(* IEC 61131-3 sources: sis-interlock-demo/tests/GVLs/Generated, 2 files *)

(* ---- GVL_TestsGenerated.gvl.st ---- *)
// AUTO-GENERATED by cemgen 1.0.0 — не редактировать: правьте матрицу и запустите
//   python -m cemgen generate <файл матрицы .csv или .xlsx>
// Матрица: SIS-V101-CEM, объект V-101, ревизия B от 2026-10-19, SHA-256 сетки df2ed4841a9453ca
// Назначение: экземпляры сгенерированных наборов coUnit: таблицы истинности голосования и сценарии
//             по матрице. {attribute 'linkalways'} обязателен: без него CODESYS выбрасывает GVL, на
//             которую никто не ссылается, и наборы молча пропадают.
// Автор:      kr0nsch; код — генератор cemgen
// Версия:     1.0.0
// Документ:   docs/DESIGN.md, раздел «10. Генератор cemgen»; docs/cause_effect_matrix.md
// ВНИМАНИЕ:   код демонстрационный и не предназначен для систем безопасности. Реальная ПАЗ требует
//             определения SIL, сертифицированных аппаратных и программных средств и валидации по
//             ГОСТ Р МЭК 61511.
{attribute 'qualified_only'}
{attribute 'linkalways'}
VAR_GLOBAL
    fbVoteTruthTest : FB_VoteTruth_Test;   // таблицы истинности голосования (36 тестов)
    fbCemGen01Test  : FB_CemGen01_Test;    // сценарии по матрице, тесты 1–40
    fbCemGen02Test  : FB_CemGen02_Test;    // сценарии по матрице, тесты 41–80
    fbCemGen03Test  : FB_CemGen03_Test;    // сценарии по матрице, тесты 81–83
END_VAR

(* ---- GVL_VoteTruthTable.gvl.st ---- *)
// AUTO-GENERATED by cemgen 1.0.0 — не редактировать: правьте матрицу и запустите
//   python -m cemgen generate <файл матрицы .csv или .xlsx>
// Матрица: SIS-V101-CEM, объект V-101, ревизия B от 2026-10-19, SHA-256 сетки df2ed4841a9453ca
// Назначение: таблицы истинности голосования (DESIGN.md, 12.2): ожидаемые байты результата
//             F_VoteEval (уровень 1) и FB_Voting (уровень 2) для всех схем, политик и видов входа;
//             считает эталонная модель cemgen. Байт: бит 0 — xTrip, бит 1 — xDegraded, биты 2–4 —
//             eArchEff (0 None, 1 1oo1, 2 1oo2, 3 2oo2, 4 2oo3, 5 ForcedTrip), биты 5–7 — байпас
//             каналов 1–3 Active (уровень 2).
// Автор:      kr0nsch; код — генератор cemgen
// Версия:     1.0.0
// Документ:   docs/DESIGN.md, раздел «10. Генератор cemgen»; docs/cause_effect_matrix.md
// ВНИМАНИЕ:   код демонстрационный и не предназначен для систем безопасности. Реальная ПАЗ требует
//             определения SIL, сертифицированных аппаратных и программных средств и валидации по
//             ГОСТ Р МЭК 61511.
{attribute 'qualified_only'}
VAR_GLOBAL CONSTANT
    // Уровень 1 — F_VoteEval: строка r, состояние канала k — (r SHR 2(k − 1)) AND 3:
    // 0 Normal, 1 Demand, 2 Invalid, 3 Bypassed; каналы k > N — NotUsed
    TT_EVAL_1OO1_VT : ARRAY[0..3] OF BYTE := [
        16#04, 16#05, 16#17, 16#17];
    TT_EVAL_1OO1_DS : ARRAY[0..3] OF BYTE := [
        16#04, 16#05, 16#17, 16#17];
    TT_EVAL_1OO1_DA : ARRAY[0..3] OF BYTE := [
        16#04, 16#05, 16#17, 16#17];
    TT_EVAL_1OO2_VT : ARRAY[0..15] OF BYTE := [
        16#08, 16#09, 16#17, 16#06, 16#09, 16#09, 16#17, 16#07, 16#17, 16#17, 16#17, 16#17, 16#06, 16#07, 16#17, 16#17];
    TT_EVAL_1OO2_DS : ARRAY[0..15] OF BYTE := [
        16#08, 16#09, 16#06, 16#06, 16#09, 16#09, 16#07, 16#07, 16#06, 16#07, 16#17, 16#17, 16#06, 16#07, 16#17, 16#17];
    TT_EVAL_1OO2_DA : ARRAY[0..15] OF BYTE := [
        16#08, 16#09, 16#06, 16#06, 16#09, 16#09, 16#07, 16#07, 16#06, 16#07, 16#17, 16#17, 16#06, 16#07, 16#17, 16#17];
    TT_EVAL_2OO2_VT : ARRAY[0..15] OF BYTE := [
        16#0C, 16#0C, 16#06, 16#06, 16#0C, 16#0D, 16#07, 16#07, 16#06, 16#07, 16#17, 16#17, 16#06, 16#07, 16#17, 16#17];
    TT_EVAL_2OO2_DS : ARRAY[0..15] OF BYTE := [
        16#0C, 16#0C, 16#06, 16#06, 16#0C, 16#0D, 16#07, 16#07, 16#06, 16#07, 16#17, 16#17, 16#06, 16#07, 16#17, 16#17];
    TT_EVAL_2OO2_DA : ARRAY[0..15] OF BYTE := [
        16#0C, 16#0C, 16#06, 16#06, 16#0C, 16#0D, 16#07, 16#07, 16#06, 16#07, 16#17, 16#17, 16#06, 16#07, 16#17, 16#17];
    TT_EVAL_2OO3_VT : ARRAY[0..63] OF BYTE := [
        16#10, 16#10, 16#0A, 16#0A, 16#10, 16#11, 16#0B, 16#0B, 16#0A, 16#0B, 16#17, 16#17, 16#0A, 16#0B, 16#17, 16#06,
        16#10, 16#11, 16#0B, 16#0B, 16#11, 16#11, 16#0B, 16#0B, 16#0B, 16#0B, 16#17, 16#17, 16#0B, 16#0B, 16#17, 16#07,
        16#0A, 16#0B, 16#17, 16#17, 16#0B, 16#0B, 16#17, 16#17, 16#17, 16#17, 16#17, 16#17, 16#17, 16#17, 16#17, 16#17,
        16#0A, 16#0B, 16#17, 16#06, 16#0B, 16#0B, 16#17, 16#07, 16#17, 16#17, 16#17, 16#17, 16#06, 16#07, 16#17, 16#17];
    TT_EVAL_2OO3_DS : ARRAY[0..63] OF BYTE := [
        16#10, 16#10, 16#0A, 16#0A, 16#10, 16#11, 16#0B, 16#0B, 16#0A, 16#0B, 16#06, 16#06, 16#0A, 16#0B, 16#06, 16#06,
        16#10, 16#11, 16#0B, 16#0B, 16#11, 16#11, 16#0B, 16#0B, 16#0B, 16#0B, 16#07, 16#07, 16#0B, 16#0B, 16#07, 16#07,
        16#0A, 16#0B, 16#06, 16#06, 16#0B, 16#0B, 16#07, 16#07, 16#06, 16#07, 16#17, 16#17, 16#06, 16#07, 16#17, 16#17,
        16#0A, 16#0B, 16#06, 16#06, 16#0B, 16#0B, 16#07, 16#07, 16#06, 16#07, 16#17, 16#17, 16#06, 16#07, 16#17, 16#17];
    TT_EVAL_2OO3_DA : ARRAY[0..63] OF BYTE := [
        16#10, 16#10, 16#0E, 16#0E, 16#10, 16#11, 16#0E, 16#0E, 16#0E, 16#0E, 16#06, 16#06, 16#0E, 16#0E, 16#06, 16#06,
        16#10, 16#11, 16#0E, 16#0E, 16#11, 16#11, 16#0F, 16#0F, 16#0E, 16#0F, 16#07, 16#07, 16#0E, 16#0F, 16#07, 16#07,
        16#0E, 16#0E, 16#06, 16#06, 16#0E, 16#0F, 16#07, 16#07, 16#06, 16#07, 16#17, 16#17, 16#06, 16#07, 16#17, 16#17,
        16#0E, 16#0E, 16#06, 16#06, 16#0E, 16#0F, 16#07, 16#07, 16#06, 16#07, 16#17, 16#17, 16#06, 16#07, 16#17, 16#17];
    // Уровень 2 — FB_Voting: строка r, биты канала k — 3(k − 1): требование, достоверность,
    // запрос байпаса; на строку два вызова одного экземпляра (сначала без запросов байпаса)
    TT_FB_1OO1_VT_DI : ARRAY[0..7] OF BYTE := [
        16#17, 16#17, 16#04, 16#05, 16#17, 16#17, 16#04, 16#05];
    TT_FB_1OO1_VT_AI : ARRAY[0..7] OF BYTE := [
        16#17, 16#17, 16#04, 16#05, 16#17, 16#17, 16#04, 16#05];
    TT_FB_1OO1_DS_DI : ARRAY[0..7] OF BYTE := [
        16#17, 16#17, 16#04, 16#05, 16#17, 16#17, 16#04, 16#05];
    TT_FB_1OO1_DS_AI : ARRAY[0..7] OF BYTE := [
        16#17, 16#17, 16#04, 16#05, 16#17, 16#17, 16#04, 16#05];
    TT_FB_1OO1_DA_DI : ARRAY[0..7] OF BYTE := [
        16#17, 16#17, 16#04, 16#05, 16#17, 16#17, 16#04, 16#05];
    TT_FB_1OO1_DA_AI : ARRAY[0..7] OF BYTE := [
        16#17, 16#17, 16#04, 16#05, 16#17, 16#17, 16#04, 16#05];
    TT_FB_1OO2_VT_DI : ARRAY[0..63] OF BYTE := [
        16#17, 16#17, 16#17, 16#17, 16#37, 16#37, 16#37, 16#37, 16#17, 16#17, 16#17, 16#17, 16#37, 16#37, 16#37, 16#37,
        16#17, 16#17, 16#08, 16#09, 16#26, 16#26, 16#26, 16#26, 16#17, 16#17, 16#09, 16#09, 16#27, 16#27, 16#27, 16#27,
        16#57, 16#57, 16#46, 16#47, 16#37, 16#37, 16#37, 16#37, 16#57, 16#57, 16#46, 16#47, 16#37, 16#37, 16#37, 16#37,
        16#57, 16#57, 16#46, 16#47, 16#26, 16#26, 16#26, 16#26, 16#57, 16#57, 16#46, 16#47, 16#27, 16#27, 16#27, 16#27];
    TT_FB_1OO2_VT_AI : ARRAY[0..63] OF BYTE := [
        16#17, 16#17, 16#17, 16#17, 16#37, 16#37, 16#37, 16#37, 16#17, 16#17, 16#17, 16#17, 16#37, 16#37, 16#37, 16#37,
        16#17, 16#17, 16#08, 16#09, 16#26, 16#26, 16#26, 16#26, 16#17, 16#17, 16#09, 16#09, 16#27, 16#27, 16#27, 16#27,
        16#57, 16#57, 16#46, 16#47, 16#37, 16#37, 16#37, 16#37, 16#57, 16#57, 16#46, 16#47, 16#37, 16#37, 16#37, 16#37,
        16#57, 16#57, 16#46, 16#47, 16#26, 16#26, 16#26, 16#26, 16#57, 16#57, 16#46, 16#47, 16#27, 16#27, 16#27, 16#27];
    TT_FB_1OO2_DS_DI : ARRAY[0..63] OF BYTE := [
        16#17, 16#17, 16#06, 16#07, 16#37, 16#37, 16#37, 16#37, 16#17, 16#17, 16#06, 16#07, 16#37, 16#37, 16#37, 16#37,
        16#06, 16#06, 16#08, 16#09, 16#26, 16#26, 16#26, 16#26, 16#07, 16#07, 16#09, 16#09, 16#27, 16#27, 16#27, 16#27,
        16#57, 16#57, 16#46, 16#47, 16#37, 16#37, 16#37, 16#37, 16#57, 16#57, 16#46, 16#47, 16#37, 16#37, 16#37, 16#37,
        16#57, 16#57, 16#46, 16#47, 16#26, 16#26, 16#26, 16#26, 16#57, 16#57, 16#46, 16#47, 16#27, 16#27, 16#27, 16#27];
    TT_FB_1OO2_DS_AI : ARRAY[0..63] OF BYTE := [
        16#17, 16#17, 16#06, 16#07, 16#37, 16#37, 16#37, 16#37, 16#17, 16#17, 16#06, 16#07, 16#37, 16#37, 16#37, 16#37,
        16#06, 16#06, 16#08, 16#09, 16#26, 16#26, 16#26, 16#26, 16#07, 16#07, 16#09, 16#09, 16#27, 16#27, 16#27, 16#27,
        16#57, 16#57, 16#46, 16#47, 16#37, 16#37, 16#37, 16#37, 16#57, 16#57, 16#46, 16#47, 16#37, 16#37, 16#37, 16#37,
        16#57, 16#57, 16#46, 16#47, 16#26, 16#26, 16#26, 16#26, 16#57, 16#57, 16#46, 16#47, 16#27, 16#27, 16#27, 16#27];
    TT_FB_1OO2_DA_DI : ARRAY[0..63] OF BYTE := [
        16#17, 16#17, 16#06, 16#07, 16#37, 16#37, 16#37, 16#37, 16#17, 16#17, 16#06, 16#07, 16#37, 16#37, 16#37, 16#37,
        16#06, 16#06, 16#08, 16#09, 16#26, 16#26, 16#26, 16#26, 16#07, 16#07, 16#09, 16#09, 16#27, 16#27, 16#27, 16#27,
        16#57, 16#57, 16#46, 16#47, 16#37, 16#37, 16#37, 16#37, 16#57, 16#57, 16#46, 16#47, 16#37, 16#37, 16#37, 16#37,
        16#57, 16#57, 16#46, 16#47, 16#26, 16#26, 16#26, 16#26, 16#57, 16#57, 16#46, 16#47, 16#27, 16#27, 16#27, 16#27];
    TT_FB_1OO2_DA_AI : ARRAY[0..63] OF BYTE := [
        16#17, 16#17, 16#06, 16#07, 16#37, 16#37, 16#37, 16#37, 16#17, 16#17, 16#06, 16#07, 16#37, 16#37, 16#37, 16#37,
        16#06, 16#06, 16#08, 16#09, 16#26, 16#26, 16#26, 16#26, 16#07, 16#07, 16#09, 16#09, 16#27, 16#27, 16#27, 16#27,
        16#57, 16#57, 16#46, 16#47, 16#37, 16#37, 16#37, 16#37, 16#57, 16#57, 16#46, 16#47, 16#37, 16#37, 16#37, 16#37,
        16#57, 16#57, 16#46, 16#47, 16#26, 16#26, 16#26, 16#26, 16#57, 16#57, 16#46, 16#47, 16#27, 16#27, 16#27, 16#27];
    TT_FB_2OO2_VT_DI : ARRAY[0..63] OF BYTE := [
        16#17, 16#17, 16#06, 16#07, 16#37, 16#37, 16#37, 16#37, 16#17, 16#17, 16#06, 16#07, 16#37, 16#37, 16#37, 16#37,
        16#06, 16#06, 16#0C, 16#0C, 16#26, 16#26, 16#26, 16#26, 16#07, 16#07, 16#0C, 16#0D, 16#27, 16#27, 16#27, 16#27,
        16#57, 16#57, 16#46, 16#47, 16#37, 16#37, 16#37, 16#37, 16#57, 16#57, 16#46, 16#47, 16#37, 16#37, 16#37, 16#37,
        16#57, 16#57, 16#46, 16#47, 16#26, 16#26, 16#26, 16#26, 16#57, 16#57, 16#46, 16#47, 16#27, 16#27, 16#27, 16#27];
    TT_FB_2OO2_VT_AI : ARRAY[0..63] OF BYTE := [
        16#17, 16#17, 16#06, 16#07, 16#37, 16#37, 16#37, 16#37, 16#17, 16#17, 16#06, 16#07, 16#37, 16#37, 16#37, 16#37,
        16#06, 16#06, 16#0C, 16#0C, 16#26, 16#26, 16#26, 16#26, 16#07, 16#07, 16#0C, 16#0D, 16#27, 16#27, 16#27, 16#27,
        16#57, 16#57, 16#46, 16#47, 16#37, 16#37, 16#37, 16#37, 16#57, 16#57, 16#46, 16#47, 16#37, 16#37, 16#37, 16#37,
        16#57, 16#57, 16#46, 16#47, 16#26, 16#26, 16#26, 16#26, 16#57, 16#57, 16#46, 16#47, 16#27, 16#27, 16#27, 16#27];
    TT_FB_2OO2_DS_DI : ARRAY[0..63] OF BYTE := [
        16#17, 16#17, 16#06, 16#07, 16#37, 16#37, 16#37, 16#37, 16#17, 16#17, 16#06, 16#07, 16#37, 16#37, 16#37, 16#37,
        16#06, 16#06, 16#0C, 16#0C, 16#26, 16#26, 16#26, 16#26, 16#07, 16#07, 16#0C, 16#0D, 16#27, 16#27, 16#27, 16#27,
        16#57, 16#57, 16#46, 16#47, 16#37, 16#37, 16#37, 16#37, 16#57, 16#57, 16#46, 16#47, 16#37, 16#37, 16#37, 16#37,
        16#57, 16#57, 16#46, 16#47, 16#26, 16#26, 16#26, 16#26, 16#57, 16#57, 16#46, 16#47, 16#27, 16#27, 16#27, 16#27];
    TT_FB_2OO2_DS_AI : ARRAY[0..63] OF BYTE := [
        16#17, 16#17, 16#06, 16#07, 16#37, 16#37, 16#37, 16#37, 16#17, 16#17, 16#06, 16#07, 16#37, 16#37, 16#37, 16#37,
        16#06, 16#06, 16#0C, 16#0C, 16#26, 16#26, 16#26, 16#26, 16#07, 16#07, 16#0C, 16#0D, 16#27, 16#27, 16#27, 16#27,
        16#57, 16#57, 16#46, 16#47, 16#37, 16#37, 16#37, 16#37, 16#57, 16#57, 16#46, 16#47, 16#37, 16#37, 16#37, 16#37,
        16#57, 16#57, 16#46, 16#47, 16#26, 16#26, 16#26, 16#26, 16#57, 16#57, 16#46, 16#47, 16#27, 16#27, 16#27, 16#27];
    TT_FB_2OO2_DA_DI : ARRAY[0..63] OF BYTE := [
        16#17, 16#17, 16#06, 16#07, 16#37, 16#37, 16#37, 16#37, 16#17, 16#17, 16#06, 16#07, 16#37, 16#37, 16#37, 16#37,
        16#06, 16#06, 16#0C, 16#0C, 16#26, 16#26, 16#26, 16#26, 16#07, 16#07, 16#0C, 16#0D, 16#27, 16#27, 16#27, 16#27,
        16#57, 16#57, 16#46, 16#47, 16#37, 16#37, 16#37, 16#37, 16#57, 16#57, 16#46, 16#47, 16#37, 16#37, 16#37, 16#37,
        16#57, 16#57, 16#46, 16#47, 16#26, 16#26, 16#26, 16#26, 16#57, 16#57, 16#46, 16#47, 16#27, 16#27, 16#27, 16#27];
    TT_FB_2OO2_DA_AI : ARRAY[0..63] OF BYTE := [
        16#17, 16#17, 16#06, 16#07, 16#37, 16#37, 16#37, 16#37, 16#17, 16#17, 16#06, 16#07, 16#37, 16#37, 16#37, 16#37,
        16#06, 16#06, 16#0C, 16#0C, 16#26, 16#26, 16#26, 16#26, 16#07, 16#07, 16#0C, 16#0D, 16#27, 16#27, 16#27, 16#27,
        16#57, 16#57, 16#46, 16#47, 16#37, 16#37, 16#37, 16#37, 16#57, 16#57, 16#46, 16#47, 16#37, 16#37, 16#37, 16#37,
        16#57, 16#57, 16#46, 16#47, 16#26, 16#26, 16#26, 16#26, 16#57, 16#57, 16#46, 16#47, 16#27, 16#27, 16#27, 16#27];
    TT_FB_2OO3_VT_DI : ARRAY[0..511] OF BYTE := [
        16#17, 16#17, 16#17, 16#17, 16#37, 16#37, 16#37, 16#37, 16#17, 16#17, 16#17, 16#17, 16#37, 16#37, 16#37, 16#37,
        16#17, 16#17, 16#0A, 16#0B, 16#37, 16#37, 16#37, 16#37, 16#17, 16#17, 16#0B, 16#0B, 16#37, 16#37, 16#37, 16#37,
        16#57, 16#57, 16#57, 16#57, 16#37, 16#37, 16#37, 16#37, 16#57, 16#57, 16#57, 16#57, 16#37, 16#37, 16#37, 16#37,
        16#57, 16#57, 16#57, 16#57, 16#37, 16#37, 16#37, 16#37, 16#57, 16#57, 16#57, 16#57, 16#37, 16#37, 16#37, 16#37,
        16#17, 16#17, 16#17, 16#17, 16#37, 16#37, 16#37, 16#37, 16#17, 16#17, 16#17, 16#17, 16#37, 16#37, 16#37, 16#37,
        16#17, 16#17, 16#0A, 16#0B, 16#37, 16#37, 16#37, 16#37, 16#17, 16#17, 16#0B, 16#0B, 16#37, 16#37, 16#37, 16#37,
        16#57, 16#57, 16#57, 16#57, 16#37, 16#37, 16#37, 16#37, 16#57, 16#57, 16#57, 16#57, 16#37, 16#37, 16#37, 16#37,
        16#57, 16#57, 16#57, 16#57, 16#37, 16#37, 16#37, 16#37, 16#57, 16#57, 16#57, 16#57, 16#37, 16#37, 16#37, 16#37,
        16#17, 16#17, 16#0A, 16#0B, 16#37, 16#37, 16#37, 16#37, 16#17, 16#17, 16#0A, 16#0B, 16#37, 16#37, 16#37, 16#37,
        16#0A, 16#0A, 16#10, 16#10, 16#2A, 16#2A, 16#2A, 16#2A, 16#0B, 16#0B, 16#10, 16#11, 16#2B, 16#2B, 16#2B, 16#2B,
        16#57, 16#57, 16#4A, 16#4B, 16#37, 16#37, 16#37, 16#37, 16#57, 16#57, 16#4A, 16#4B, 16#37, 16#37, 16#37, 16#37,
        16#57, 16#57, 16#4A, 16#4B, 16#2A, 16#2A, 16#2A, 16#2A, 16#57, 16#57, 16#4A, 16#4B, 16#2B, 16#2B, 16#2B, 16#2B,
        16#17, 16#17, 16#0B, 16#0B, 16#37, 16#37, 16#37, 16#37, 16#17, 16#17, 16#0B, 16#0B, 16#37, 16#37, 16#37, 16#37,
        16#0B, 16#0B, 16#10, 16#11, 16#2B, 16#2B, 16#2B, 16#2B, 16#0B, 16#0B, 16#11, 16#11, 16#2B, 16#2B, 16#2B, 16#2B,
        16#57, 16#57, 16#4B, 16#4B, 16#37, 16#37, 16#37, 16#37, 16#57, 16#57, 16#4B, 16#4B, 16#37, 16#37, 16#37, 16#37,
        16#57, 16#57, 16#4B, 16#4B, 16#2B, 16#2B, 16#2B, 16#2B, 16#57, 16#57, 16#4B, 16#4B, 16#2B, 16#2B, 16#2B, 16#2B,
        16#97, 16#97, 16#97, 16#97, 16#37, 16#37, 16#37, 16#37, 16#97, 16#97, 16#97, 16#97, 16#37, 16#37, 16#37, 16#37,
        16#97, 16#97, 16#8A, 16#8B, 16#37, 16#37, 16#37, 16#37, 16#97, 16#97, 16#8B, 16#8B, 16#37, 16#37, 16#37, 16#37,
        16#57, 16#57, 16#57, 16#57, 16#37, 16#37, 16#37, 16#37, 16#57, 16#57, 16#57, 16#57, 16#37, 16#37, 16#37, 16#37,
        16#57, 16#57, 16#57, 16#57, 16#37, 16#37, 16#37, 16#37, 16#57, 16#57, 16#57, 16#57, 16#37, 16#37, 16#37, 16#37,
        16#97, 16#97, 16#97, 16#97, 16#37, 16#37, 16#37, 16#37, 16#97, 16#97, 16#97, 16#97, 16#37, 16#37, 16#37, 16#37,
        16#97, 16#97, 16#8A, 16#8B, 16#37, 16#37, 16#37, 16#37, 16#97, 16#97, 16#8B, 16#8B, 16#37, 16#37, 16#37, 16#37,
        16#57, 16#57, 16#57, 16#57, 16#37, 16#37, 16#37, 16#37, 16#57, 16#57, 16#57, 16#57, 16#37, 16#37, 16#37, 16#37,
        16#57, 16#57, 16#57, 16#57, 16#37, 16#37, 16#37, 16#37, 16#57, 16#57, 16#57, 16#57, 16#37, 16#37, 16#37, 16#37,
        16#97, 16#97, 16#97, 16#97, 16#37, 16#37, 16#37, 16#37, 16#97, 16#97, 16#97, 16#97, 16#37, 16#37, 16#37, 16#37,
        16#97, 16#97, 16#8A, 16#8B, 16#2A, 16#2A, 16#2A, 16#2A, 16#97, 16#97, 16#8B, 16#8B, 16#2B, 16#2B, 16#2B, 16#2B,
        16#57, 16#57, 16#4A, 16#4B, 16#37, 16#37, 16#37, 16#37, 16#57, 16#57, 16#4A, 16#4B, 16#37, 16#37, 16#37, 16#37,
        16#57, 16#57, 16#4A, 16#4B, 16#2A, 16#2A, 16#2A, 16#2A, 16#57, 16#57, 16#4A, 16#4B, 16#2B, 16#2B, 16#2B, 16#2B,
        16#97, 16#97, 16#97, 16#97, 16#37, 16#37, 16#37, 16#37, 16#97, 16#97, 16#97, 16#97, 16#37, 16#37, 16#37, 16#37,
        16#97, 16#97, 16#8A, 16#8B, 16#2B, 16#2B, 16#2B, 16#2B, 16#97, 16#97, 16#8B, 16#8B, 16#2B, 16#2B, 16#2B, 16#2B,
        16#57, 16#57, 16#4B, 16#4B, 16#37, 16#37, 16#37, 16#37, 16#57, 16#57, 16#4B, 16#4B, 16#37, 16#37, 16#37, 16#37,
        16#57, 16#57, 16#4B, 16#4B, 16#2B, 16#2B, 16#2B, 16#2B, 16#57, 16#57, 16#4B, 16#4B, 16#2B, 16#2B, 16#2B, 16#2B];
    TT_FB_2OO3_VT_AI : ARRAY[0..511] OF BYTE := [
        16#17, 16#17, 16#17, 16#17, 16#37, 16#37, 16#37, 16#37, 16#17, 16#17, 16#17, 16#17, 16#37, 16#37, 16#37, 16#37,
        16#17, 16#17, 16#0A, 16#0B, 16#37, 16#37, 16#37, 16#37, 16#17, 16#17, 16#0B, 16#0B, 16#37, 16#37, 16#37, 16#37,
        16#57, 16#57, 16#57, 16#57, 16#37, 16#37, 16#37, 16#37, 16#57, 16#57, 16#57, 16#57, 16#37, 16#37, 16#37, 16#37,
        16#57, 16#57, 16#57, 16#57, 16#37, 16#37, 16#37, 16#37, 16#57, 16#57, 16#57, 16#57, 16#37, 16#37, 16#37, 16#37,
        16#17, 16#17, 16#17, 16#17, 16#37, 16#37, 16#37, 16#37, 16#17, 16#17, 16#17, 16#17, 16#37, 16#37, 16#37, 16#37,
        16#17, 16#17, 16#0A, 16#0B, 16#37, 16#37, 16#37, 16#37, 16#17, 16#17, 16#0B, 16#0B, 16#37, 16#37, 16#37, 16#37,
        16#57, 16#57, 16#57, 16#57, 16#37, 16#37, 16#37, 16#37, 16#57, 16#57, 16#57, 16#57, 16#37, 16#37, 16#37, 16#37,
        16#57, 16#57, 16#57, 16#57, 16#37, 16#37, 16#37, 16#37, 16#57, 16#57, 16#57, 16#57, 16#37, 16#37, 16#37, 16#37,
        16#17, 16#17, 16#0A, 16#0B, 16#37, 16#37, 16#37, 16#37, 16#17, 16#17, 16#0A, 16#0B, 16#37, 16#37, 16#37, 16#37,
        16#0A, 16#0A, 16#10, 16#10, 16#2A, 16#2A, 16#2A, 16#2A, 16#0B, 16#0B, 16#10, 16#11, 16#2B, 16#2B, 16#2B, 16#2B,
        16#57, 16#57, 16#4A, 16#4B, 16#37, 16#37, 16#37, 16#37, 16#57, 16#57, 16#4A, 16#4B, 16#37, 16#37, 16#37, 16#37,
        16#57, 16#57, 16#4A, 16#4B, 16#2A, 16#2A, 16#2A, 16#2A, 16#57, 16#57, 16#4A, 16#4B, 16#2B, 16#2B, 16#2B, 16#2B,
        16#17, 16#17, 16#0B, 16#0B, 16#37, 16#37, 16#37, 16#37, 16#17, 16#17, 16#0B, 16#0B, 16#37, 16#37, 16#37, 16#37,
        16#0B, 16#0B, 16#10, 16#11, 16#2B, 16#2B, 16#2B, 16#2B, 16#0B, 16#0B, 16#11, 16#11, 16#2B, 16#2B, 16#2B, 16#2B,
        16#57, 16#57, 16#4B, 16#4B, 16#37, 16#37, 16#37, 16#37, 16#57, 16#57, 16#4B, 16#4B, 16#37, 16#37, 16#37, 16#37,
        16#57, 16#57, 16#4B, 16#4B, 16#2B, 16#2B, 16#2B, 16#2B, 16#57, 16#57, 16#4B, 16#4B, 16#2B, 16#2B, 16#2B, 16#2B,
        16#97, 16#97, 16#97, 16#97, 16#37, 16#37, 16#37, 16#37, 16#97, 16#97, 16#97, 16#97, 16#37, 16#37, 16#37, 16#37,
        16#97, 16#97, 16#8A, 16#8B, 16#37, 16#37, 16#37, 16#37, 16#97, 16#97, 16#8B, 16#8B, 16#37, 16#37, 16#37, 16#37,
        16#57, 16#57, 16#57, 16#57, 16#37, 16#37, 16#37, 16#37, 16#57, 16#57, 16#57, 16#57, 16#37, 16#37, 16#37, 16#37,
        16#57, 16#57, 16#57, 16#57, 16#37, 16#37, 16#37, 16#37, 16#57, 16#57, 16#57, 16#57, 16#37, 16#37, 16#37, 16#37,
        16#97, 16#97, 16#97, 16#97, 16#37, 16#37, 16#37, 16#37, 16#97, 16#97, 16#97, 16#97, 16#37, 16#37, 16#37, 16#37,
        16#97, 16#97, 16#8A, 16#8B, 16#37, 16#37, 16#37, 16#37, 16#97, 16#97, 16#8B, 16#8B, 16#37, 16#37, 16#37, 16#37,
        16#57, 16#57, 16#57, 16#57, 16#37, 16#37, 16#37, 16#37, 16#57, 16#57, 16#57, 16#57, 16#37, 16#37, 16#37, 16#37,
        16#57, 16#57, 16#57, 16#57, 16#37, 16#37, 16#37, 16#37, 16#57, 16#57, 16#57, 16#57, 16#37, 16#37, 16#37, 16#37,
        16#97, 16#97, 16#97, 16#97, 16#37, 16#37, 16#37, 16#37, 16#97, 16#97, 16#97, 16#97, 16#37, 16#37, 16#37, 16#37,
        16#97, 16#97, 16#8A, 16#8B, 16#2A, 16#2A, 16#2A, 16#2A, 16#97, 16#97, 16#8B, 16#8B, 16#2B, 16#2B, 16#2B, 16#2B,
        16#57, 16#57, 16#4A, 16#4B, 16#37, 16#37, 16#37, 16#37, 16#57, 16#57, 16#4A, 16#4B, 16#37, 16#37, 16#37, 16#37,
        16#57, 16#57, 16#4A, 16#4B, 16#2A, 16#2A, 16#2A, 16#2A, 16#57, 16#57, 16#4A, 16#4B, 16#2B, 16#2B, 16#2B, 16#2B,
        16#97, 16#97, 16#97, 16#97, 16#37, 16#37, 16#37, 16#37, 16#97, 16#97, 16#97, 16#97, 16#37, 16#37, 16#37, 16#37,
        16#97, 16#97, 16#8A, 16#8B, 16#2B, 16#2B, 16#2B, 16#2B, 16#97, 16#97, 16#8B, 16#8B, 16#2B, 16#2B, 16#2B, 16#2B,
        16#57, 16#57, 16#4B, 16#4B, 16#37, 16#37, 16#37, 16#37, 16#57, 16#57, 16#4B, 16#4B, 16#37, 16#37, 16#37, 16#37,
        16#57, 16#57, 16#4B, 16#4B, 16#2B, 16#2B, 16#2B, 16#2B, 16#57, 16#57, 16#4B, 16#4B, 16#2B, 16#2B, 16#2B, 16#2B];
    TT_FB_2OO3_DS_DI : ARRAY[0..511] OF BYTE := [
        16#17, 16#17, 16#06, 16#07, 16#37, 16#37, 16#37, 16#37, 16#17, 16#17, 16#06, 16#07, 16#37, 16#37, 16#37, 16#37,
        16#06, 16#06, 16#0A, 16#0B, 16#26, 16#26, 16#26, 16#26, 16#07, 16#07, 16#0B, 16#0B, 16#27, 16#27, 16#27, 16#27,
        16#57, 16#57, 16#46, 16#47, 16#37, 16#37, 16#37, 16#37, 16#57, 16#57, 16#46, 16#47, 16#37, 16#37, 16#37, 16#37,
        16#57, 16#57, 16#46, 16#47, 16#26, 16#26, 16#26, 16#26, 16#57, 16#57, 16#46, 16#47, 16#27, 16#27, 16#27, 16#27,
        16#17, 16#17, 16#06, 16#07, 16#37, 16#37, 16#37, 16#37, 16#17, 16#17, 16#06, 16#07, 16#37, 16#37, 16#37, 16#37,
        16#06, 16#06, 16#0A, 16#0B, 16#26, 16#26, 16#26, 16#26, 16#07, 16#07, 16#0B, 16#0B, 16#27, 16#27, 16#27, 16#27,
        16#57, 16#57, 16#46, 16#47, 16#37, 16#37, 16#37, 16#37, 16#57, 16#57, 16#46, 16#47, 16#37, 16#37, 16#37, 16#37,
        16#57, 16#57, 16#46, 16#47, 16#26, 16#26, 16#26, 16#26, 16#57, 16#57, 16#46, 16#47, 16#27, 16#27, 16#27, 16#27,
        16#06, 16#06, 16#0A, 16#0B, 16#26, 16#26, 16#26, 16#26, 16#06, 16#06, 16#0A, 16#0B, 16#26, 16#26, 16#26, 16#26,
        16#0A, 16#0A, 16#10, 16#10, 16#2A, 16#2A, 16#2A, 16#2A, 16#0B, 16#0B, 16#10, 16#11, 16#2B, 16#2B, 16#2B, 16#2B,
        16#46, 16#46, 16#4A, 16#4B, 16#26, 16#26, 16#26, 16#26, 16#46, 16#46, 16#4A, 16#4B, 16#26, 16#26, 16#26, 16#26,
        16#46, 16#46, 16#4A, 16#4B, 16#2A, 16#2A, 16#2A, 16#2A, 16#46, 16#46, 16#4A, 16#4B, 16#2B, 16#2B, 16#2B, 16#2B,
        16#07, 16#07, 16#0B, 16#0B, 16#27, 16#27, 16#27, 16#27, 16#07, 16#07, 16#0B, 16#0B, 16#27, 16#27, 16#27, 16#27,
        16#0B, 16#0B, 16#10, 16#11, 16#2B, 16#2B, 16#2B, 16#2B, 16#0B, 16#0B, 16#11, 16#11, 16#2B, 16#2B, 16#2B, 16#2B,
        16#47, 16#47, 16#4B, 16#4B, 16#27, 16#27, 16#27, 16#27, 16#47, 16#47, 16#4B, 16#4B, 16#27, 16#27, 16#27, 16#27,
        16#47, 16#47, 16#4B, 16#4B, 16#2B, 16#2B, 16#2B, 16#2B, 16#47, 16#47, 16#4B, 16#4B, 16#2B, 16#2B, 16#2B, 16#2B,
        16#97, 16#97, 16#86, 16#87, 16#37, 16#37, 16#37, 16#37, 16#97, 16#97, 16#86, 16#87, 16#37, 16#37, 16#37, 16#37,
        16#86, 16#86, 16#8A, 16#8B, 16#26, 16#26, 16#26, 16#26, 16#87, 16#87, 16#8B, 16#8B, 16#27, 16#27, 16#27, 16#27,
        16#57, 16#57, 16#46, 16#47, 16#37, 16#37, 16#37, 16#37, 16#57, 16#57, 16#46, 16#47, 16#37, 16#37, 16#37, 16#37,
        16#57, 16#57, 16#46, 16#47, 16#26, 16#26, 16#26, 16#26, 16#57, 16#57, 16#46, 16#47, 16#27, 16#27, 16#27, 16#27,
        16#97, 16#97, 16#86, 16#87, 16#37, 16#37, 16#37, 16#37, 16#97, 16#97, 16#86, 16#87, 16#37, 16#37, 16#37, 16#37,
        16#86, 16#86, 16#8A, 16#8B, 16#26, 16#26, 16#26, 16#26, 16#87, 16#87, 16#8B, 16#8B, 16#27, 16#27, 16#27, 16#27,
        16#57, 16#57, 16#46, 16#47, 16#37, 16#37, 16#37, 16#37, 16#57, 16#57, 16#46, 16#47, 16#37, 16#37, 16#37, 16#37,
        16#57, 16#57, 16#46, 16#47, 16#26, 16#26, 16#26, 16#26, 16#57, 16#57, 16#46, 16#47, 16#27, 16#27, 16#27, 16#27,
        16#97, 16#97, 16#86, 16#87, 16#26, 16#26, 16#26, 16#26, 16#97, 16#97, 16#86, 16#87, 16#26, 16#26, 16#26, 16#26,
        16#86, 16#86, 16#8A, 16#8B, 16#2A, 16#2A, 16#2A, 16#2A, 16#87, 16#87, 16#8B, 16#8B, 16#2B, 16#2B, 16#2B, 16#2B,
        16#46, 16#46, 16#4A, 16#4B, 16#26, 16#26, 16#26, 16#26, 16#46, 16#46, 16#4A, 16#4B, 16#26, 16#26, 16#26, 16#26,
        16#46, 16#46, 16#4A, 16#4B, 16#2A, 16#2A, 16#2A, 16#2A, 16#46, 16#46, 16#4A, 16#4B, 16#2B, 16#2B, 16#2B, 16#2B,
        16#97, 16#97, 16#86, 16#87, 16#27, 16#27, 16#27, 16#27, 16#97, 16#97, 16#86, 16#87, 16#27, 16#27, 16#27, 16#27,
        16#86, 16#86, 16#8A, 16#8B, 16#2B, 16#2B, 16#2B, 16#2B, 16#87, 16#87, 16#8B, 16#8B, 16#2B, 16#2B, 16#2B, 16#2B,
        16#47, 16#47, 16#4B, 16#4B, 16#27, 16#27, 16#27, 16#27, 16#47, 16#47, 16#4B, 16#4B, 16#27, 16#27, 16#27, 16#27,
        16#47, 16#47, 16#4B, 16#4B, 16#2B, 16#2B, 16#2B, 16#2B, 16#47, 16#47, 16#4B, 16#4B, 16#2B, 16#2B, 16#2B, 16#2B];
    TT_FB_2OO3_DS_AI : ARRAY[0..511] OF BYTE := [
        16#17, 16#17, 16#06, 16#07, 16#37, 16#37, 16#37, 16#37, 16#17, 16#17, 16#06, 16#07, 16#37, 16#37, 16#37, 16#37,
        16#06, 16#06, 16#0A, 16#0B, 16#26, 16#26, 16#26, 16#26, 16#07, 16#07, 16#0B, 16#0B, 16#27, 16#27, 16#27, 16#27,
        16#57, 16#57, 16#46, 16#47, 16#37, 16#37, 16#37, 16#37, 16#57, 16#57, 16#46, 16#47, 16#37, 16#37, 16#37, 16#37,
        16#57, 16#57, 16#46, 16#47, 16#26, 16#26, 16#26, 16#26, 16#57, 16#57, 16#46, 16#47, 16#27, 16#27, 16#27, 16#27,
        16#17, 16#17, 16#06, 16#07, 16#37, 16#37, 16#37, 16#37, 16#17, 16#17, 16#06, 16#07, 16#37, 16#37, 16#37, 16#37,
        16#06, 16#06, 16#0A, 16#0B, 16#26, 16#26, 16#26, 16#26, 16#07, 16#07, 16#0B, 16#0B, 16#27, 16#27, 16#27, 16#27,
        16#57, 16#57, 16#46, 16#47, 16#37, 16#37, 16#37, 16#37, 16#57, 16#57, 16#46, 16#47, 16#37, 16#37, 16#37, 16#37,
        16#57, 16#57, 16#46, 16#47, 16#26, 16#26, 16#26, 16#26, 16#57, 16#57, 16#46, 16#47, 16#27, 16#27, 16#27, 16#27,
        16#06, 16#06, 16#0A, 16#0B, 16#26, 16#26, 16#26, 16#26, 16#06, 16#06, 16#0A, 16#0B, 16#26, 16#26, 16#26, 16#26,
        16#0A, 16#0A, 16#10, 16#10, 16#2A, 16#2A, 16#2A, 16#2A, 16#0B, 16#0B, 16#10, 16#11, 16#2B, 16#2B, 16#2B, 16#2B,
        16#46, 16#46, 16#4A, 16#4B, 16#26, 16#26, 16#26, 16#26, 16#46, 16#46, 16#4A, 16#4B, 16#26, 16#26, 16#26, 16#26,
        16#46, 16#46, 16#4A, 16#4B, 16#2A, 16#2A, 16#2A, 16#2A, 16#46, 16#46, 16#4A, 16#4B, 16#2B, 16#2B, 16#2B, 16#2B,
        16#07, 16#07, 16#0B, 16#0B, 16#27, 16#27, 16#27, 16#27, 16#07, 16#07, 16#0B, 16#0B, 16#27, 16#27, 16#27, 16#27,
        16#0B, 16#0B, 16#10, 16#11, 16#2B, 16#2B, 16#2B, 16#2B, 16#0B, 16#0B, 16#11, 16#11, 16#2B, 16#2B, 16#2B, 16#2B,
        16#47, 16#47, 16#4B, 16#4B, 16#27, 16#27, 16#27, 16#27, 16#47, 16#47, 16#4B, 16#4B, 16#27, 16#27, 16#27, 16#27,
        16#47, 16#47, 16#4B, 16#4B, 16#2B, 16#2B, 16#2B, 16#2B, 16#47, 16#47, 16#4B, 16#4B, 16#2B, 16#2B, 16#2B, 16#2B,
        16#97, 16#97, 16#86, 16#87, 16#37, 16#37, 16#37, 16#37, 16#97, 16#97, 16#86, 16#87, 16#37, 16#37, 16#37, 16#37,
        16#86, 16#86, 16#8A, 16#8B, 16#26, 16#26, 16#26, 16#26, 16#87, 16#87, 16#8B, 16#8B, 16#27, 16#27, 16#27, 16#27,
        16#57, 16#57, 16#46, 16#47, 16#37, 16#37, 16#37, 16#37, 16#57, 16#57, 16#46, 16#47, 16#37, 16#37, 16#37, 16#37,
        16#57, 16#57, 16#46, 16#47, 16#26, 16#26, 16#26, 16#26, 16#57, 16#57, 16#46, 16#47, 16#27, 16#27, 16#27, 16#27,
        16#97, 16#97, 16#86, 16#87, 16#37, 16#37, 16#37, 16#37, 16#97, 16#97, 16#86, 16#87, 16#37, 16#37, 16#37, 16#37,
        16#86, 16#86, 16#8A, 16#8B, 16#26, 16#26, 16#26, 16#26, 16#87, 16#87, 16#8B, 16#8B, 16#27, 16#27, 16#27, 16#27,
        16#57, 16#57, 16#46, 16#47, 16#37, 16#37, 16#37, 16#37, 16#57, 16#57, 16#46, 16#47, 16#37, 16#37, 16#37, 16#37,
        16#57, 16#57, 16#46, 16#47, 16#26, 16#26, 16#26, 16#26, 16#57, 16#57, 16#46, 16#47, 16#27, 16#27, 16#27, 16#27,
        16#97, 16#97, 16#86, 16#87, 16#26, 16#26, 16#26, 16#26, 16#97, 16#97, 16#86, 16#87, 16#26, 16#26, 16#26, 16#26,
        16#86, 16#86, 16#8A, 16#8B, 16#2A, 16#2A, 16#2A, 16#2A, 16#87, 16#87, 16#8B, 16#8B, 16#2B, 16#2B, 16#2B, 16#2B,
        16#46, 16#46, 16#4A, 16#4B, 16#26, 16#26, 16#26, 16#26, 16#46, 16#46, 16#4A, 16#4B, 16#26, 16#26, 16#26, 16#26,
        16#46, 16#46, 16#4A, 16#4B, 16#2A, 16#2A, 16#2A, 16#2A, 16#46, 16#46, 16#4A, 16#4B, 16#2B, 16#2B, 16#2B, 16#2B,
        16#97, 16#97, 16#86, 16#87, 16#27, 16#27, 16#27, 16#27, 16#97, 16#97, 16#86, 16#87, 16#27, 16#27, 16#27, 16#27,
        16#86, 16#86, 16#8A, 16#8B, 16#2B, 16#2B, 16#2B, 16#2B, 16#87, 16#87, 16#8B, 16#8B, 16#2B, 16#2B, 16#2B, 16#2B,
        16#47, 16#47, 16#4B, 16#4B, 16#27, 16#27, 16#27, 16#27, 16#47, 16#47, 16#4B, 16#4B, 16#27, 16#27, 16#27, 16#27,
        16#47, 16#47, 16#4B, 16#4B, 16#2B, 16#2B, 16#2B, 16#2B, 16#47, 16#47, 16#4B, 16#4B, 16#2B, 16#2B, 16#2B, 16#2B];
    TT_FB_2OO3_DA_DI : ARRAY[0..511] OF BYTE := [
        16#17, 16#17, 16#06, 16#07, 16#37, 16#37, 16#37, 16#37, 16#17, 16#17, 16#06, 16#07, 16#37, 16#37, 16#37, 16#37,
        16#06, 16#06, 16#0E, 16#0E, 16#26, 16#26, 16#26, 16#26, 16#07, 16#07, 16#0E, 16#0F, 16#27, 16#27, 16#27, 16#27,
        16#57, 16#57, 16#46, 16#47, 16#37, 16#37, 16#37, 16#37, 16#57, 16#57, 16#46, 16#47, 16#37, 16#37, 16#37, 16#37,
        16#57, 16#57, 16#46, 16#47, 16#26, 16#26, 16#26, 16#26, 16#57, 16#57, 16#46, 16#47, 16#27, 16#27, 16#27, 16#27,
        16#17, 16#17, 16#06, 16#07, 16#37, 16#37, 16#37, 16#37, 16#17, 16#17, 16#06, 16#07, 16#37, 16#37, 16#37, 16#37,
        16#06, 16#06, 16#0E, 16#0E, 16#26, 16#26, 16#26, 16#26, 16#07, 16#07, 16#0E, 16#0F, 16#27, 16#27, 16#27, 16#27,
        16#57, 16#57, 16#46, 16#47, 16#37, 16#37, 16#37, 16#37, 16#57, 16#57, 16#46, 16#47, 16#37, 16#37, 16#37, 16#37,
        16#57, 16#57, 16#46, 16#47, 16#26, 16#26, 16#26, 16#26, 16#57, 16#57, 16#46, 16#47, 16#27, 16#27, 16#27, 16#27,
        16#06, 16#06, 16#0E, 16#0E, 16#26, 16#26, 16#26, 16#26, 16#06, 16#06, 16#0E, 16#0E, 16#26, 16#26, 16#26, 16#26,
        16#0E, 16#0E, 16#10, 16#10, 16#2E, 16#2E, 16#2E, 16#2E, 16#0E, 16#0E, 16#10, 16#11, 16#2E, 16#2E, 16#2E, 16#2E,
        16#46, 16#46, 16#4E, 16#4E, 16#26, 16#26, 16#26, 16#26, 16#46, 16#46, 16#4E, 16#4E, 16#26, 16#26, 16#26, 16#26,
        16#46, 16#46, 16#4E, 16#4E, 16#2E, 16#2E, 16#2E, 16#2E, 16#46, 16#46, 16#4E, 16#4E, 16#2E, 16#2E, 16#2E, 16#2E,
        16#07, 16#07, 16#0E, 16#0F, 16#27, 16#27, 16#27, 16#27, 16#07, 16#07, 16#0E, 16#0F, 16#27, 16#27, 16#27, 16#27,
        16#0E, 16#0E, 16#10, 16#11, 16#2E, 16#2E, 16#2E, 16#2E, 16#0F, 16#0F, 16#11, 16#11, 16#2F, 16#2F, 16#2F, 16#2F,
        16#47, 16#47, 16#4E, 16#4F, 16#27, 16#27, 16#27, 16#27, 16#47, 16#47, 16#4E, 16#4F, 16#27, 16#27, 16#27, 16#27,
        16#47, 16#47, 16#4E, 16#4F, 16#2E, 16#2E, 16#2E, 16#2E, 16#47, 16#47, 16#4E, 16#4F, 16#2F, 16#2F, 16#2F, 16#2F,
        16#97, 16#97, 16#86, 16#87, 16#37, 16#37, 16#37, 16#37, 16#97, 16#97, 16#86, 16#87, 16#37, 16#37, 16#37, 16#37,
        16#86, 16#86, 16#8E, 16#8E, 16#26, 16#26, 16#26, 16#26, 16#87, 16#87, 16#8E, 16#8F, 16#27, 16#27, 16#27, 16#27,
        16#57, 16#57, 16#46, 16#47, 16#37, 16#37, 16#37, 16#37, 16#57, 16#57, 16#46, 16#47, 16#37, 16#37, 16#37, 16#37,
        16#57, 16#57, 16#46, 16#47, 16#26, 16#26, 16#26, 16#26, 16#57, 16#57, 16#46, 16#47, 16#27, 16#27, 16#27, 16#27,
        16#97, 16#97, 16#86, 16#87, 16#37, 16#37, 16#37, 16#37, 16#97, 16#97, 16#86, 16#87, 16#37, 16#37, 16#37, 16#37,
        16#86, 16#86, 16#8E, 16#8E, 16#26, 16#26, 16#26, 16#26, 16#87, 16#87, 16#8E, 16#8F, 16#27, 16#27, 16#27, 16#27,
        16#57, 16#57, 16#46, 16#47, 16#37, 16#37, 16#37, 16#37, 16#57, 16#57, 16#46, 16#47, 16#37, 16#37, 16#37, 16#37,
        16#57, 16#57, 16#46, 16#47, 16#26, 16#26, 16#26, 16#26, 16#57, 16#57, 16#46, 16#47, 16#27, 16#27, 16#27, 16#27,
        16#97, 16#97, 16#86, 16#87, 16#26, 16#26, 16#26, 16#26, 16#97, 16#97, 16#86, 16#87, 16#26, 16#26, 16#26, 16#26,
        16#86, 16#86, 16#8E, 16#8E, 16#2E, 16#2E, 16#2E, 16#2E, 16#87, 16#87, 16#8E, 16#8F, 16#2E, 16#2E, 16#2E, 16#2E,
        16#46, 16#46, 16#4E, 16#4E, 16#26, 16#26, 16#26, 16#26, 16#46, 16#46, 16#4E, 16#4E, 16#26, 16#26, 16#26, 16#26,
        16#46, 16#46, 16#4E, 16#4E, 16#2E, 16#2E, 16#2E, 16#2E, 16#46, 16#46, 16#4E, 16#4E, 16#2E, 16#2E, 16#2E, 16#2E,
        16#97, 16#97, 16#86, 16#87, 16#27, 16#27, 16#27, 16#27, 16#97, 16#97, 16#86, 16#87, 16#27, 16#27, 16#27, 16#27,
        16#86, 16#86, 16#8E, 16#8E, 16#2E, 16#2E, 16#2E, 16#2E, 16#87, 16#87, 16#8E, 16#8F, 16#2F, 16#2F, 16#2F, 16#2F,
        16#47, 16#47, 16#4E, 16#4F, 16#27, 16#27, 16#27, 16#27, 16#47, 16#47, 16#4E, 16#4F, 16#27, 16#27, 16#27, 16#27,
        16#47, 16#47, 16#4E, 16#4F, 16#2E, 16#2E, 16#2E, 16#2E, 16#47, 16#47, 16#4E, 16#4F, 16#2F, 16#2F, 16#2F, 16#2F];
    TT_FB_2OO3_DA_AI : ARRAY[0..511] OF BYTE := [
        16#17, 16#17, 16#06, 16#07, 16#37, 16#37, 16#37, 16#37, 16#17, 16#17, 16#06, 16#07, 16#37, 16#37, 16#37, 16#37,
        16#06, 16#06, 16#0E, 16#0E, 16#26, 16#26, 16#26, 16#26, 16#07, 16#07, 16#0E, 16#0F, 16#27, 16#27, 16#27, 16#27,
        16#57, 16#57, 16#46, 16#47, 16#37, 16#37, 16#37, 16#37, 16#57, 16#57, 16#46, 16#47, 16#37, 16#37, 16#37, 16#37,
        16#57, 16#57, 16#46, 16#47, 16#26, 16#26, 16#26, 16#26, 16#57, 16#57, 16#46, 16#47, 16#27, 16#27, 16#27, 16#27,
        16#17, 16#17, 16#06, 16#07, 16#37, 16#37, 16#37, 16#37, 16#17, 16#17, 16#06, 16#07, 16#37, 16#37, 16#37, 16#37,
        16#06, 16#06, 16#0E, 16#0E, 16#26, 16#26, 16#26, 16#26, 16#07, 16#07, 16#0E, 16#0F, 16#27, 16#27, 16#27, 16#27,
        16#57, 16#57, 16#46, 16#47, 16#37, 16#37, 16#37, 16#37, 16#57, 16#57, 16#46, 16#47, 16#37, 16#37, 16#37, 16#37,
        16#57, 16#57, 16#46, 16#47, 16#26, 16#26, 16#26, 16#26, 16#57, 16#57, 16#46, 16#47, 16#27, 16#27, 16#27, 16#27,
        16#06, 16#06, 16#0E, 16#0E, 16#26, 16#26, 16#26, 16#26, 16#06, 16#06, 16#0E, 16#0E, 16#26, 16#26, 16#26, 16#26,
        16#0E, 16#0E, 16#10, 16#10, 16#2E, 16#2E, 16#2E, 16#2E, 16#0E, 16#0E, 16#10, 16#11, 16#2E, 16#2E, 16#2E, 16#2E,
        16#46, 16#46, 16#4E, 16#4E, 16#26, 16#26, 16#26, 16#26, 16#46, 16#46, 16#4E, 16#4E, 16#26, 16#26, 16#26, 16#26,
        16#46, 16#46, 16#4E, 16#4E, 16#2E, 16#2E, 16#2E, 16#2E, 16#46, 16#46, 16#4E, 16#4E, 16#2E, 16#2E, 16#2E, 16#2E,
        16#07, 16#07, 16#0E, 16#0F, 16#27, 16#27, 16#27, 16#27, 16#07, 16#07, 16#0E, 16#0F, 16#27, 16#27, 16#27, 16#27,
        16#0E, 16#0E, 16#10, 16#11, 16#2E, 16#2E, 16#2E, 16#2E, 16#0F, 16#0F, 16#11, 16#11, 16#2F, 16#2F, 16#2F, 16#2F,
        16#47, 16#47, 16#4E, 16#4F, 16#27, 16#27, 16#27, 16#27, 16#47, 16#47, 16#4E, 16#4F, 16#27, 16#27, 16#27, 16#27,
        16#47, 16#47, 16#4E, 16#4F, 16#2E, 16#2E, 16#2E, 16#2E, 16#47, 16#47, 16#4E, 16#4F, 16#2F, 16#2F, 16#2F, 16#2F,
        16#97, 16#97, 16#86, 16#87, 16#37, 16#37, 16#37, 16#37, 16#97, 16#97, 16#86, 16#87, 16#37, 16#37, 16#37, 16#37,
        16#86, 16#86, 16#8E, 16#8E, 16#26, 16#26, 16#26, 16#26, 16#87, 16#87, 16#8E, 16#8F, 16#27, 16#27, 16#27, 16#27,
        16#57, 16#57, 16#46, 16#47, 16#37, 16#37, 16#37, 16#37, 16#57, 16#57, 16#46, 16#47, 16#37, 16#37, 16#37, 16#37,
        16#57, 16#57, 16#46, 16#47, 16#26, 16#26, 16#26, 16#26, 16#57, 16#57, 16#46, 16#47, 16#27, 16#27, 16#27, 16#27,
        16#97, 16#97, 16#86, 16#87, 16#37, 16#37, 16#37, 16#37, 16#97, 16#97, 16#86, 16#87, 16#37, 16#37, 16#37, 16#37,
        16#86, 16#86, 16#8E, 16#8E, 16#26, 16#26, 16#26, 16#26, 16#87, 16#87, 16#8E, 16#8F, 16#27, 16#27, 16#27, 16#27,
        16#57, 16#57, 16#46, 16#47, 16#37, 16#37, 16#37, 16#37, 16#57, 16#57, 16#46, 16#47, 16#37, 16#37, 16#37, 16#37,
        16#57, 16#57, 16#46, 16#47, 16#26, 16#26, 16#26, 16#26, 16#57, 16#57, 16#46, 16#47, 16#27, 16#27, 16#27, 16#27,
        16#97, 16#97, 16#86, 16#87, 16#26, 16#26, 16#26, 16#26, 16#97, 16#97, 16#86, 16#87, 16#26, 16#26, 16#26, 16#26,
        16#86, 16#86, 16#8E, 16#8E, 16#2E, 16#2E, 16#2E, 16#2E, 16#87, 16#87, 16#8E, 16#8F, 16#2E, 16#2E, 16#2E, 16#2E,
        16#46, 16#46, 16#4E, 16#4E, 16#26, 16#26, 16#26, 16#26, 16#46, 16#46, 16#4E, 16#4E, 16#26, 16#26, 16#26, 16#26,
        16#46, 16#46, 16#4E, 16#4E, 16#2E, 16#2E, 16#2E, 16#2E, 16#46, 16#46, 16#4E, 16#4E, 16#2E, 16#2E, 16#2E, 16#2E,
        16#97, 16#97, 16#86, 16#87, 16#27, 16#27, 16#27, 16#27, 16#97, 16#97, 16#86, 16#87, 16#27, 16#27, 16#27, 16#27,
        16#86, 16#86, 16#8E, 16#8E, 16#2E, 16#2E, 16#2E, 16#2E, 16#87, 16#87, 16#8E, 16#8F, 16#2F, 16#2F, 16#2F, 16#2F,
        16#47, 16#47, 16#4E, 16#4F, 16#27, 16#27, 16#27, 16#27, 16#47, 16#47, 16#4E, 16#4F, 16#27, 16#27, 16#27, 16#27,
        16#47, 16#47, 16#4E, 16#4F, 16#2E, 16#2E, 16#2E, 16#2E, 16#47, 16#47, 16#4E, 16#4F, 16#2F, 16#2F, 16#2F, 16#2F];
END_VAR
